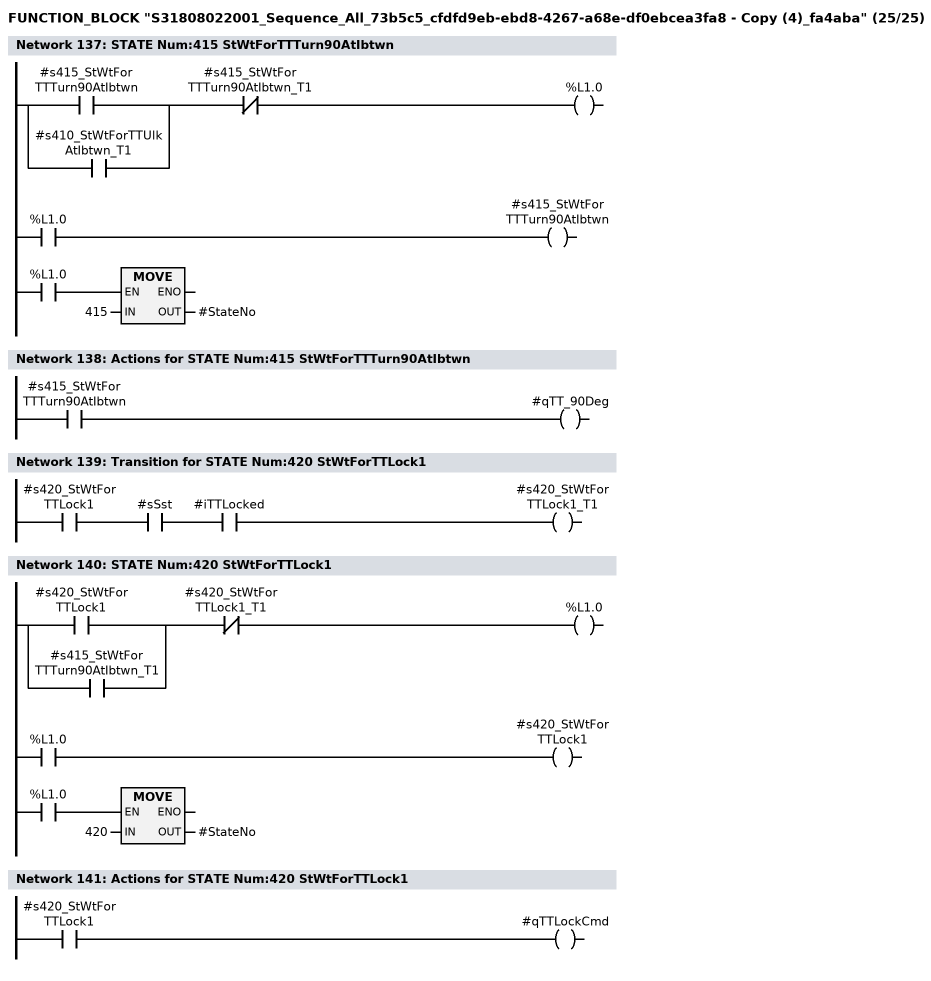
      A(;
      O #s415_StWtForTTTurn90AtIbtwn;
      O #s410_StWtForTTUlkAtIbtwn_T1;
      );
      AN #s415_StWtForTTTurn90AtIbtwn_T1;
      = %L1.0;
      A %L1.0;
      BLD 102;
      = #s415_StWtForTTTurn90AtIbtwn;
      A %L1.0;
      JNB Label_415;
      L 415;
      T #StateNo;
Label_415:      NOP 0;
NETWORK
TITLE = Actions for STATE Num:415 StWtForTTTurn90AtIbtwn
      A #s415_StWtForTTTurn90AtIbtwn;
      = #qTT_90Deg;
NETWORK
TITLE = Transition for STATE Num:420 StWtForTTLock1
      A #s420_StWtForTTLock1;
      A #sSst;
      A #iTTLocked;
      = #s420_StWtForTTLock1_T1;
NETWORK
TITLE = STATE Num:420 StWtForTTLock1
      A(;
      O #s420_StWtForTTLock1;
      O #s415_StWtForTTTurn90AtIbtwn_T1;
      );
      AN #s420_StWtForTTLock1_T1;
      = %L1.0;
      A %L1.0;
      BLD 102;
      = #s420_StWtForTTLock1;
      A %L1.0;
      JNB Label_420;
      L 420;
      T #StateNo;
Label_420:      NOP 0;
NETWORK
TITLE = Actions for STATE Num:420 StWtForTTLock1
      A #s420_StWtForTTLock1;
      = #qTTLockCmd;
END_FUNCTION_BLOCK